FUNCTION_BLOCK TypeScopeTest (* Basic FB validating current type lookup *)
  (* Standard: 61499-1; Description: Copyright (c) 2026 Martin Erich Jobst This program and the accompanying materials are made available under the terms of the Eclipse Public License 2.0 which is available at https://www.eclipse.org/legal/epl-2.0/ SPDX-License-Identifier: EPL-2.0 *)
  (* Version 1.0, 2026-11-18, Martin Jobst *)
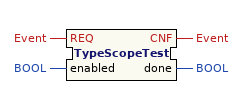
  EVENT_INPUT
    REQ; (* Request *)
  END_EVENT
  EVENT_OUTPUT
    CNF; (* Confirmation *)
  END_EVENT
  VAR_INPUT
    enabled : BOOL := TRUE;
  END_VAR
  VAR_OUTPUT
    done : BOOL := initialState;
  END_VAR
  VAR CONSTANT
    initialState : BOOL := TRUE;
  END_VAR
  VAR
    state : BOOL := initialState;
  END_VAR
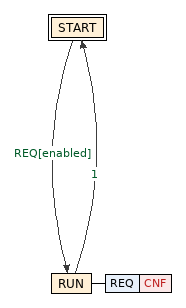
  EC_STATES
    START;
    RUN : REQ -> CNF;
  END_STATES
  EC_TRANSITIONS
    START TO RUN := REQ[enabled];
    RUN TO START := 1;
  END_TRANSITIONS
  ALGORITHM REQ IN ST:
state := enabled;
done := state;
  END_ALGORITHM
END_FUNCTION_BLOCK
